Staubli VAL3: physicalIO.pgx

program physicalIO()
// Level 3: four taught piston slots with tool presence sensing and bounded assembly.
begin
  // ============================================================
  // SENSORES Y ALIMENTADOR DEL LEVEL 3
  // ============================================================
  // Solo se crea en fisico. En simulacion los sensores se editan a mano.
  // La pinza usa open/close con valve1; NO escribir valve1 aqui.
  while true
    pistonPresent = io:bIn0 == true
    cylinderPresent = io:bIn2 == true
    feederExtended = io:bIn14 == true
    feederRetracted = io:bIn15 == true
    io:bOut10 = feederExtend
    ioReady = true
    delay(0.01)
  endWhile
end
